Staubli VAL3: initImage.pgx

public program initImage(utImage& x_utImage[], string x_sPage, string x_sId)
begin
  x_utImage.Common.sPage=x_sPage
  x_utImage.Common.sID=x_sId
  userPageBind(x_utImage.Common.sPage,x_utImage.Common.sID,"src",x_utImage.Common.sSourceImage,1,"r")
  userPageBind(x_utImage.Common.sPage,x_utImage.Common.sID,"style.visibility",x_utImage.Appearance.bVisibility,1,"r")
  userPageBindClick(x_utImage.Common.sPage,x_utImage.Common.sID,x_utImage.Events.bClick,true)
  //
  userPageBind(x_utImage.Common.sPage,x_utImage.Common.sID,"className",x_utImage.Common.sClass,1,"r")
  //userPageBind(x_sPage,x_utImage.Common.sID,"style.borderColor",x_utImage.Border.sBorderColour,1,"r")
  //userPageBind(x_sPage,x_utImage.Common.sID,"style.borderStyle",x_utImage.Border.sBorderStyle,1,"r")
  //
  x_utImage.Appearance.bVisibility=true
  x_utImage.Events.bClick=false
  x_utImage.Common.sClass="clickable"
end
